Fanuc KAREL source: KT00509.KL

PROGRAM KT00509
%NOLOCKGROUP
VAR
  P1: XYZWPR
  P2: JOINTPOS
  OUT: POSITION
BEGIN
  P1.X = 1.0
  OUT = P1 : P2
END KT00509
